(* IEC 61131-3 sources: codesys-to-astra/cds2astra/tests/corpus/C2A-RET001/pos/src/GVLs, 1 file *)

(* ---- GVL_R.gvl.st ---- *)
// Назначение: корпус правила cds2astra (synthetic).
// Автор:      kr0nsch
// Версия:     0.1.0
// Документ:   docs/RULES.md
VAR_GLOBAL RETAIN
    udiCnt : UDINT; // счётчик
END_VAR
